(* IEC 61131-3 sources: llm-plc-st-eval/data/raw/claude-sonnet-4-6/B1/zero_shot, 3 files *)

(* ---- ejec_1.st ---- *)
```pascal
FUNCTION_BLOCK FB_Motor
VAR_INPUT
    btnMarcha : BOOL; (* Botón de marcha: TRUE = pulsado *)
    btnParo   : BOOL; (* Botón de paro: TRUE = pulsado *)
    btnEmerg  : BOOL; (* Paro de emergencia: TRUE = activado *)
END_VAR

VAR_OUTPUT
    motorOn : BOOL; (* Salida al contactor del motor *)
END_VAR

VAR
    bloqueado : BOOL; (* Enclavamiento por emergencia *)
END_VAR

(*
    Lógica de control:
    1. Si se activa la emergencia → parar motor y bloquear rearranque.
    2. El bloqueo se mantiene mientras btnEmerg siga activo.
    3. Si se pulsa paro → apagar motor (sin bloqueo).
    4. Si se pulsa marcha y no hay bloqueo → encender motor (auto-retención).
*)

(* --- Gestión del enclavamiento de emergencia --- *)
IF btnEmerg THEN
    bloqueado := TRUE;   (* Activar bloqueo *)
    motorOn   := FALSE;  (* Parar motor inmediatamente *)
ELSIF NOT btnEmerg THEN
    bloqueado := FALSE;  (* Liberar bloqueo cuando se rearma la emergencia *)
END_IF;

(* --- Lógica de marcha / paro (solo si no hay bloqueo) --- *)
IF NOT bloqueado THEN
    IF btnParo THEN
        motorOn := FALSE; (* Paro normal *)
    ELSIF btnMarcha THEN
        motorOn := TRUE;  (* Arranque con auto-retención *)
    END_IF;
END_IF;

END_FUNCTION_BLOCK
```

(* ---- ejec_2.st ---- *)
```pascal
FUNCTION_BLOCK FB_Motor
VAR_INPUT
    btnMarcha : BOOL; (* Botón de marcha: TRUE = pulsado *)
    btnParo   : BOOL; (* Botón de paro: TRUE = pulsado *)
    btnEmerg  : BOOL; (* Paro de emergencia: TRUE = activado *)
END_VAR

VAR_OUTPUT
    motorOn : BOOL; (* Salida al contactor del motor *)
END_VAR

VAR
    bloqueEmerg : BOOL := FALSE; (* Enclavamiento por emergencia *)
END_VAR

(*
    Lógica de control:
    1. Si se activa la emergencia: parar motor y bloquear rearranque.
    2. El bloqueo de emergencia solo se libera cuando btnEmerg vuelve
       a FALSE (rearme manual implícito al soltar la seta).
    3. Si no hay bloqueo: SET con btnMarcha, RESET con btnParo.
*)

(* --- Gestión del enclavamiento de emergencia --- *)
IF btnEmerg THEN
    bloqueEmerg := TRUE;  (* Activar bloqueo *)
ELSIF NOT btnEmerg THEN
    bloqueEmerg := FALSE; (* Liberar bloqueo al soltar la seta *)
END_IF;

(* --- Lógica de marcha / paro con enclavamiento --- *)
IF bloqueEmerg OR btnParo THEN
    (* Paro prioritario: emergencia o botón de paro *)
    motorOn := FALSE;
ELSIF btnMarcha AND NOT bloqueEmerg THEN
    (* Arranque: solo si no hay bloqueo activo *)
    motorOn := TRUE;
END_IF;
(* Si ninguna condición aplica, motorOn conserva su valor anterior
   (efecto de memoria / auto-mantenimiento). *)

END_FUNCTION_BLOCK
```

(* ---- ejec_3.st ---- *)
```pascal
FUNCTION_BLOCK FB_Motor
VAR_INPUT
    btnMarcha : BOOL; (* Botón de marcha: TRUE = pulsado *)
    btnParo   : BOOL; (* Botón de paro: TRUE = pulsado *)
    btnEmerg  : BOOL; (* Paro de emergencia: TRUE = activado *)
END_VAR

VAR_OUTPUT
    motorOn : BOOL; (* Salida al contactor del motor *)
END_VAR

VAR
    bloqueEmerg : BOOL := FALSE; (* Enclavamiento por emergencia *)
END_VAR

(*
    Lógica de control:
    1. Si se activa la emergencia → parar motor y bloquear rearranque.
    2. El bloqueo de emergencia solo se libera cuando btnEmerg vuelve
       a FALSE (emergencia restablecida) Y el botón de marcha NO está
       pulsado, evitando un arranque automático no deseado.
    3. Paro normal → apaga el motor sin bloqueo.
    4. Marcha → arranca solo si no hay bloqueo activo.
    5. Autoretención: motorOn se mantiene mientras no haya paro.
*)

(* --- Gestión del enclavamiento de emergencia --- *)
IF btnEmerg THEN
    (* Emergencia activa: bloquear y apagar *)
    bloqueEmerg := TRUE;
    motorOn     := FALSE;

ELSIF bloqueEmerg THEN
    (* Emergencia ya restablecida (btnEmerg = FALSE):
       liberar bloqueo solo si el botón de marcha no está pulsado *)
    IF NOT btnMarcha THEN
        bloqueEmerg := FALSE;
    END_IF;
    motorOn := FALSE; (* Motor permanece parado mientras haya bloqueo *)

ELSE
    (* Funcionamiento normal: sin emergencia ni bloqueo *)

    IF btnParo THEN
        (* Paro normal: apagar motor *)
        motorOn := FALSE;

    ELSIF btnMarcha THEN
        (* Arranque: activar motor *)
        motorOn := TRUE;

    END_IF;
    (* Si ningún botón está pulsado, motorOn conserva su valor → autoretención *)

END_IF;
```
